PROGRAM PRG_Lamp
VAR
	bLamp	: BOOL;
END_VAR

END_PROGRAM

(* stored: Version 1.1.0.1
   POU PRG_Lamp: Id {aae628a3-c8a7-4043-b338-7b14460910c8}, SpecialFunc None *)
